Fanuc KAREL source: compact_preamble.KL

PROGRAM KB00088
%NOLOCKGROUP
VAR
P1:INTEGER;P2:INTEGER;P3:INTEGER;RESULT : XYZWPREXT
BEGIN
P1=1
P2=1
P3=1
RESULT=GET_POS_TPE(P1,P2,P3,1)
END KB00088
